// TIA Portal V20 export
TYPE "WT2_Kd_Status_UDT"
   STRUCT
      iHandshake : Int;
      Fehler : Struct
         bE0000_KonfigFehler : Bool;
         bE0001_Reserviert : Bool;
         bE0002_InvUngueltig : Bool;
         bE0003_Reserviert : Bool;
         bE0004_Reserviert : Bool;
         bE0005_Reserviert : Bool;
         bE0006_WasserueberdruckZuTief : Bool;
         bE0007_Reserviert : Bool;
         bE0008_Reserviert : Bool;
         bE0009_Reserviert : Bool;
         bE0010_KdPumpeFehlerBetrieb : Bool;
         bE0011_KdPumpeFehlerStillstand : Bool;
         bE0012_KonfigFehlerVdMinVerflTemp : Bool;
         b035_Reserve : Bool;
         b036_Reserve : Bool;
         b037_Reserve : Bool;
         by04_Reserve : Byte;
         by05_Reserve : Byte;
      END_STRUCT;
      Alarm : Struct
         bA1000_Reserviert : Bool;
         bA1001_SlaveAusgef : Bool;
         bA1002_Reserviert : Bool;
         bA1003_HauptMasterAusgef : Bool;
         bA1004_MKdMasterAktiv : Bool;
         bA1005_ObjektIDMehrfVorhanden : Bool;
         bA1006_Reserviert : Bool;
         bA1007_WassereingangstempZuTief : Bool;
         bA1008_AlarmNivEnschalter : Bool;
         bA1009_AlarmNiv2Endschalter : Bool;
         bA1010_Reserviert : Bool;
         bA1011_Reserviert : Bool;
         bA1012_Reserviert : Bool;
         b075_Reserve : Bool;
         b076_Reserve : Bool;
         b077_Reserve : Bool;
         by08_Reserve : Byte;
         by09_Reserve : Byte;
      END_STRUCT;
      Zustand : Struct
         bFehlerzustandAktiv : Bool;
         bAlarmzustandAktiv : Bool;
         bSystemMeldungAktiv : Bool;
         bSeviceMeldungAktiv : Bool;
         bStopManuell : Bool;
         bStopAuto : Bool;
         bStopExtern : Bool;
         bBetriebAuto : Bool;
         bBetriebManuell : Bool;
         bAnlaufAuto : Bool;
         bAnlaufManuell : Bool;
         bManuellStoppen : Bool;
         b114_Reserve : Bool;
         b115_Reserve : Bool;
         b116_Reserve : Bool;
         b117_Reserve : Bool;
         by12_Reserve : Byte;
         bInventarAufnahme : Bool;
         b131_Reserve : Bool;
         bStandbyMasterInit : Bool;
         bStandbyMasterPassiv : Bool;
         bStandbyMasterAktiv : Bool;
         bNotbetriebAktiv : Bool;
         bMasterGesperrt : Bool;
         bSollwertAnhebung : Bool;
         bKdEintrittWarm : Bool;
         b141_Reserve : Bool;
         b142_Reserve : Bool;
         b143_Reserve : Bool;
         b144_Reserve : Bool;
         b145_Reserve : Bool;
         b146_Reserve : Bool;
         b147_Reserve : Bool;
         by15_Reserve : Byte;
         by16_Reserve : Byte;
         by17_Reserve : Byte;
      END_STRUCT;
      DigIn : Struct
         b180_Reserve : Bool;
         bSollwertB : Bool;
         b182_Reserve : Bool;
         bNiveauregFreigabe : Bool;
         bNiveaureg2Freigabe : Bool;
         bWasserueberdruck : Bool;
         bNivEndschOffen : Bool;
         bNivEndschGeschl : Bool;
         bNiv2EndschOffen : Bool;
         bNiv2EndschGeschl : Bool;
         b192_Reserve : Bool;
         b193_Reserve : Bool;
         b194_Reserve : Bool;
         b195_Reserve : Bool;
         b196_Reserve : Bool;
         b197_Reserve : Bool;
         by20_Reserve : Byte;
         by21_Reserve : Byte;
      END_STRUCT;
      DigOut : Struct
         b220_Reserve : Bool;
         b221_Reserve : Bool;
         bKdPumpe : Bool;
         bNiveauregelung : Bool;
         bNiveauregelung2 : Bool;
         bNiveauregelungDO : Bool;
         bNiveauregelung2DO : Bool;
         b227_Reserve : Bool;
         by23_Reserve : Byte;
         by24_Reserve : Byte;
         by25_Reserve : Byte;
      END_STRUCT;
      chReserve1 : Char;
      chKondReglerEinheit : Char;
      rKondRegIst : Real;
      rKondRegSoll : Real;
      rKondRegOut : Real;
      iKondRegStufen : Int;
      rKondTempEintritt : Real;
      rKondTempAustritt : Real;
      rAussentemp : Real;
      rReserveReal : Array[0..1] of Real;
      byReserveByte : Array[0..1] of Byte;
   END_STRUCT;
END_TYPE
